// TIA Portal V20 export
DATA_BLOCK "Zaehler_Sicherheit_DB"   // DB203
// stored: InstanceOfName Zaehler_Sicherheit, InstanceOfType FB
"Zaehler_Sicherheit"
   // VAR RETAIN
   //    "QS_NOT-HALT_Schuetz" { S7_SetPoint := 'True'} : CTU_UDINT;
   //    "QS_NOT-HALT_Tuere_1_RST" { S7_SetPoint := 'True'} : CTU_UDINT;
   //    "QS_NOT-HALT_Tuere_1" { S7_SetPoint := 'True'} : CTU_UDINT;
   //    "QS_NOT-HALT_Tuere_2_RST" { S7_SetPoint := 'True'} : CTU_UDINT;
   //    "QS_NOT-HALT_Tuere_2" { S7_SetPoint := 'True'} : CTU_UDINT;
   //    "QS_NOT-HALT_Roboter" { S7_SetPoint := 'True'} : CTU_UDINT;
   //    QS_Sichere_Bewegung { S7_SetPoint := 'True'} : CTU_UDINT;
   //    QS_Zuhaltung_Freigeben { S7_SetPoint := 'True'} : CTU_UDINT;
   // END_VAR
BEGIN
END_DATA_BLOCK
